(* IEC 61131-3 sources: plc-process-lib/src/DUTs/Alarm, 5 files *)

(* ---- E_AlarmEventReason.dut.st ---- *)
// Назначение: причина перехода тревоги в событии ST_AlarmEvent (приёмник I_AlarmSink).
// Автор:      kr0nsch
// Версия:     0.1.0
// Документ:   docs/ARCHITECTURE.md, раздел «Тревоги»
{attribute 'qualified_only'}
{attribute 'strict'}
TYPE E_AlarmEventReason :
(
    None          := 0,
    Activated     := 1,    // условие появилось (после задержки)
    Cleared       := 2,    // условие ушло (после задержки)
    Acked         := 3,
    Shelved       := 4,
    Unshelved     := 5,    // командой
    ShelveExpired := 6,    // по таймауту
    Suppressed    := 7,
    Unsuppressed  := 8,
    OosOn         := 9,
    OosOff        := 10,
    Disabled      := 11    // тревога выключена приоритетом None: закрывающее событие
) INT;
END_TYPE

(* ---- E_AlarmPriority.dut.st ---- *)
// Назначение: приоритет тревоги. None выключает тревогу: она не формируется, событий нет.
//             Значения вне перечисления FB_Alarm считает Medium.
// Автор:      kr0nsch
// Версия:     0.1.0
// Документ:   docs/ARCHITECTURE.md, раздел «Тревоги»
{attribute 'qualified_only'}
{attribute 'strict'}
TYPE E_AlarmPriority :
(
    None     := 0,   // тревога выключена: не формируется, событий нет
    Low      := 1,
    Medium   := 2,
    High     := 3,
    Critical := 4    // резерв под аварийный уровень
) INT;
END_TYPE

(* ---- E_AlarmState.dut.st ---- *)
// Назначение: состояние тревоги по ISA-18.2: четыре базовых состояния и три наложенных
//             (по старшинству OutOfService > SuppressedByDesign > Shelved). Модель состояний —
//             сверить с ANSI/ISA-18.2-2016.
// Автор:      kr0nsch
// Версия:     0.1.0
// Документ:   docs/ARCHITECTURE.md, раздел «Тревоги»
{attribute 'qualified_only'}
{attribute 'strict'}
TYPE E_AlarmState :
(
    Normal             := 0,   // норма: условия нет, квитировано
    ActiveUnack        := 1,   // активна, не квитирована
    ActiveAck          := 2,   // активна, квитирована
    RtnUnack           := 3,   // вернулась в норму без квитирования
    Shelved            := 4,   // отложена оператором, с таймаутом
    SuppressedByDesign := 5,   // подавлена по условию (логикой)
    OutOfService       := 6    // выведена из работы вместе с устройством
) INT;
END_TYPE

(* ---- ST_AlarmCfg.dut.st ---- *)
// Назначение: параметры одной тревоги (слот astAlarm[i] в Cfg устройства). 16 байт.
//             Тип лежит в Persistent Variables приложения и заморожен в пределах 1.x (A-13).
// Автор:      kr0nsch
// Версия:     0.1.0
// Документ:   docs/ARCHITECTURE.md, раздел «Тревоги»
{attribute 'qualified_only'}
TYPE ST_AlarmCfg :
STRUCT
    ePriority  : E_AlarmPriority := E_AlarmPriority.Medium;
    tOnDelay   : TIME := T#0S;   // задержка появления
    tOffDelay  : TIME := T#0S;   // задержка снятия
    tShelveMax : TIME := T#8H;   // максимальный срок shelve; T#0S — откладывать запрещено
END_STRUCT
END_TYPE

(* ---- ST_AlarmEvent.dut.st ---- *)
// Назначение: событие перехода тревоги для приёмника I_AlarmSink (журнал приложения).
//             Астрономическое время ставит приёмник, в событии — монотонная отметка LTIME.
// Автор:      kr0nsch
// Версия:     0.1.0
// Документ:   docs/ARCHITECTURE.md, раздел «Тревоги»
{attribute 'qualified_only'}
TYPE ST_AlarmEvent :
STRUCT
    udiId     : UDINT;                // номер тревоги на объекте
    ePriority : E_AlarmPriority;
    eOldState : E_AlarmState;
    eNewState : E_AlarmState;
    eReason   : E_AlarmEventReason;
    ltTime    : LTIME;                // монотонная отметка; астрономическое время ставит приёмник
    rValue    : REAL;                 // значение процесса в момент события
END_STRUCT
END_TYPE
